{region 'Documentation'}
(*!
<summary>Uses the real scheduling algorithm with a pre-use local publisher binding.</summary>
*)
{endregion}
FUNCTION_BLOCK OrchestratorProbe EXTENDS Orchestrator

SUPER^(Task := Task);

{region 'Documentation'}
(*!
<summary>Binds isolated diagnostics before Initialize or any cyclic use.</summary>
*)
{endregion}
METHOD PUBLIC BindPublisher
VAR_INPUT
    Publisher : I_EventPublisher; //! Nonzero isolated event publisher retained before subject initialization; keep it alive through all subject use.
END_VAR
FEventPublisher := Publisher;
END_METHOD

END_FUNCTION_BLOCK

(* stored: Version 1.1.0.1
   POU OrchestratorProbe: Id {ee17f657-06fd-4006-9d66-55b7e97e6563}, SpecialFunc None
   Method BindPublisher: Id {c7a9bd2f-40ce-4de5-9850-768f57a0690f} *)
